(* IEC 61131-3 sources: plc_generation_empirical_study/datasets/_archive/pre_native_plcverif_20260810/tasks/C02_E01_basic_start_stop_latch/negative_control, 1 file *)

(* ---- NC1.st ---- *)
FUNCTION_BLOCK C02_E01_basic_start_stop_latch
VAR_INPUT
    Start : BOOL;
    Stop : BOOL;
END_VAR
VAR_OUTPUT
    Running : BOOL;
END_VAR

IF Stop THEN
    Running := FALSE;
ELSIF Start THEN
    Running := FALSE;
END_IF;

END_FUNCTION_BLOCK
